// MONET/N auxiliary sensors: mirror temperatures M1 and M2 on the EL3164 (0-10 V, ch 2 and ch 1; ch 3 is the oil
// level). Copied from MONETS's FB_MonetsTelescopeAuxiliary, which also has an M1 cell and a flange sensor that
// MONET/N does not have. Replaces HalfBROT's FB_TelescopeAuxiliary (removed, HalfBROT #21).
FUNCTION_BLOCK FB_MonetnTelescopeAuxiliary
VAR
	tempSensorM1   		AT%I*: INT;
	tempSensorM2   		AT%I*: INT;
	fbComm				: I_Comm;
	sensorM1			: MONETcommon.FB_MonetTempSensor;
	sensorM2			: MONETcommon.FB_MonetTempSensor;
END_VAR
VAR_OUTPUT
	// only valid while the matching valid flag is TRUE: a broken wire reads -50 C (MONETN#17)
	tempM1				: REAL;
	tempM2				: REAL;
	validM1				: BOOL;
	validM2				: BOOL;
END_VAR

sensorM1(iRaw := tempSensorM1, sName := 'TEMP_M1', comm := fbComm);
sensorM2(iRaw := tempSensorM2, sName := 'TEMP_M2', comm := fbComm);
tempM1 			:= sensorM1.fTemperature;
tempM2 			:= sensorM2.fTemperature;
validM1 		:= sensorM1.bValid;
validM2 		:= sensorM2.bValid;

//FB_Init is always available implicitly and it is used primarily for initialization.
//The return value is not evaluated. For a specific influence, you can also declare the
//methods explicitly and provide additional code there with the standard initialization
//code. You can evaluate the return value.
METHOD FB_Init: BOOL
VAR_INPUT
    bInitRetains	: BOOL; // TRUE: the retain variables are initialized (reset warm / reset cold)
    bInCopyCode		: BOOL;  // TRUE: the instance will be copied to the copy code afterward (online change)
	comm			: I_Comm;	   
END_VAR
THIS^.fbComm := comm;
END_METHOD

METHOD SendTelemetry : BOOL
VAR_INPUT
END_VAR
IF fbComm = 0 THEN
	RETURN;
END_IF
fbComm.PublishString('telescope', 'dome', 'AUXILIARY.SENSOR[1].NAME', 'TEMP_M1');
IF validM1 THEN
	fbComm.PublishLREAL('telescope', 'dome', 'AUXILIARY.SENSOR[1].VALUE', tempM1);
END_IF
fbComm.PublishString('telescope', 'dome', 'AUXILIARY.SENSOR[1].UNIT', 'C');
fbComm.PublishString('telescope', 'dome', 'AUXILIARY.SENSOR[2].NAME', 'TEMP_M2');
IF validM2 THEN
	fbComm.PublishLREAL('telescope', 'dome', 'AUXILIARY.SENSOR[2].VALUE', tempM2);
END_IF
fbComm.PublishString('telescope', 'dome', 'AUXILIARY.SENSOR[2].UNIT', 'C');
END_METHOD

END_FUNCTION_BLOCK

(* stored: Version 1.1.0.1, ProductVersion 3.1.4024.15
   POU FB_MonetnTelescopeAuxiliary: Id {7e31d5fd-3935-4700-ae64-3b5e25a9b947}, SpecialFunc None
   Method FB_Init: Id {34154e00-1554-42d6-b807-6241695bcfd7}
   Method SendTelemetry: Id {9e49f282-bfc0-4335-a7b7-cce199e9240a} *)
